(* IEC 61131-3 sources: STAR-PLC-Agent/results/raw/codex_matrix_resume_20261114/codex_deepseek/PUB004/generation/compiler_records/compile_01, 1 file *)

(* ---- FB_Task.st ---- *)
FUNCTION_BLOCK FB_Task
VAR_INPUT
    VISCOSITY_OK : BOOL;
    PASTE_E_STOP_NC : BOOL;
    DebounceTime : TIME;
    CycleTime : TIME;
END_VAR
VAR_OUTPUT
    VFD_RUN : BOOL := FALSE;
    PUMP_MAINT_DUE : BOOL := FALSE;
    PUMP_RUNTIME_ACC : LTIME := LTIME#0ns;
END_VAR
VAR
    debounceElapsed : TIME := TIME#0ms;
    viscosityQualified : BOOL := FALSE;
END_VAR

IF NOT PASTE_E_STOP_NC THEN
    debounceElapsed := TIME#0ms;
    viscosityQualified := FALSE;
ELSIF NOT VISCOSITY_OK THEN
    debounceElapsed := TIME#0ms;
    viscosityQualified := FALSE;
ELSE
    IF debounceElapsed >= DebounceTime THEN
        viscosityQualified := TRUE;
    END_IF;
END_IF;

VFD_RUN := PASTE_E_STOP_NC AND VISCOSITY_OK AND viscosityQualified;

IF VFD_RUN THEN
    PUMP_RUNTIME_ACC := PUMP_RUNTIME_ACC + CycleTime;
END_IF;

PUMP_MAINT_DUE := PUMP_RUNTIME_ACC >= LTIME#500h;

IF PASTE_E_STOP_NC AND VISCOSITY_OK AND NOT viscosityQualified THEN
    debounceElapsed := debounceElapsed + CycleTime;
END_IF;
END_FUNCTION_BLOCK
